# EPICS autosave request: iocBoot/iocETC/auto_settings.req
file "ETC_settings.req", P=ETC:
